Fanuc KAREL source: kx00028.KL

-- PROVISIONAL review KL for V770-1; original PC SHA256 849b9d35886d4f642747c626b39a00225ce534774a73aec12a8c1a4eedffd71f
-- Incomplete behavior may be omitted. Consult companion uncertainty JSON. Do not deploy.
PROGRAM KX00028
%NOLOCKGROUP
VAR
  I : INTEGER
  J : INTEGER
  B : BOOLEAN
  F : FILE
  S : STRING[80]
-- UNRESOLVED_DECL P type=000102
BEGIN
  -- UNRESOLVED_PC offsets 5-12; opcodes 9D,23
  -- UNRESOLVED_PC offsets 17-21; opcodes 7F
END KX00028
